Fanuc KAREL source: ko00056.KL

-- PROVISIONAL review KL for V1013-1; original PC SHA256 cb5aa1970789cefe9cc367a85be8152435168be4f16fe85eca9a788ac81fbf81
-- Incomplete behavior may be omitted. Consult companion uncertainty JSON. Do not deploy.
PROGRAM KO00056
%NOLOCKGROUP
BEGIN
  -- UNRESOLVED_PC offsets 5-12; opcodes 9D,23
  -- UNRESOLVED_PC offsets 17-69; opcodes 27,27,49,7E,AD,27,49,7E,AD,22,31,7E,4A
  -- UNRESOLVED_PC offsets 74-78; opcodes 7F
END KO00056
